(* IEC 61131-3 sources: JingjiangMoonbox/Application/Application/全局, 3 files *)

(* ---- GCL.st ---- *)
(*@CES
Name=GCL
Type=ConstantList
TypeGuid=ffbfa93a-b94d-45fc-a329-229860183b1d
Guid=bcb51df0-81a2-49d0-af31-1b6fd6cdee10
HasDeclaration=True
HasImplementation=False
*)
{DECLARATION}
VAR_GLOBAL CONSTANT
	gc_xUseNewFlyRemove: BOOL:= TRUE;(*新飞点剔除总开关:TRUE=误差平均前用KS_FlyRemove
逐帧剔除并以锁存值替换飞点,FALSE=回退旧飞点判断KS_FB_PickOutFakePoint(旧逻辑完整
保留),改后重新编译生效|Yang.zj+用于新飞点检测 2026.10.24.191149*)
	MASTER_DRIVER_TIME:REAL:= 1;(*运控周期2ms*)
//2026.1.24.215529增加月光宝盒和月光宝盒PRO的类型
	HY_YTPE_CMM_CR_PRO: WORD:= 16#6006;
	HY_YTPE_CMM_CR: WORD:= 16#6005;

	USER_MAX_STATION_NUM_V1:INT:=256;

	gc_iNum_ErrorNum_GT: INT:=3;//gt指令报错执行次数
	gc_iNum_ErrorNum_GT_LOG: INT:=300;//gt指令报错执行次数去写日志
	gc_iTime_s_ServoFailed: INT:=10;//10s伺服打开超时

	gc_lrPi: LREAL:= 3.1415926;
	MAX_UNIT_NUM: INT:=16;(*最大色组数*)
	MAX_STATION_NUM: INT:= 256;
	MAX_AXIS_NUM: INT:= 128;
	(*应对牵引周长算法增加稳速判断等待时长和模拟量滤波计算周长的时长
	默认等待10s和1s调整一次周长*)
	gc_iValueReferToLost: INT:= -32768	;										(*误差标识-丢失|*)
	gc_iValueReferToFakePoint: INT:= -32767	;									(*误差标识-飞点|*)
	gc_iValueReferToSkipTheHeader: INT:= -32766	;							(*误差标识-让料头|*)

	gc_iCycleNum_CalcGirthEvenDelay: INT:= 500;(*算周长算法稳速等待时常，推荐10s(20ms周期就是500个周期)*)
	gc_iCycleNum_CalcDelay: INT:= 500;(*周长计算间隔时长，推荐1s(20ms周期就是50个周期)*)

	gc_tmHold_PreStart				: TIME := T#3S; (* 开机预启动持续时间|该值在程序中赋值给响铃时间| 2022.5.27.143829|该值被弃用*)
	gc_tmHold_PreStart_BeiRen		: TIME := T#6s; (* 北人开机预启动持续时间|和响铃时间是分开的| 2022.5.27.143829*)
	gc_tmAlarmHold_PreStart			: TIME := T#3s; (* 开机预启动报警持续时间| *)
	GC_LRMOTORPPR					: LREAL:=4194304;//2025.7.3.175755
	gc_EXT_TSK_CYCLE_TIME		: INT := 35;(*2023.06.19.102054||niu.j||任务周期35*)
	gc_TENSION_TSK_CYCLE_TIME		: INT := 20;(*2023.06.19.102054||niu.j||任务周期35*)
	gc_MAIN_TSK_CYCLE_TIME		: INT := 10;(*2023.06.19.102054||niu.j||任务周期35*)

	MAX_CMD_NUM_PDU				: INT := 10;(* 最大pdu命令的数量 *)
	MAX_PDU_CMD_BYTES_UP		: INT := 60;(* 来源于1024/16(MAX_UNIT_NUM)/此数必须是4字节的整数倍 *)
	MAX_PDU_CMD_BYTES_DN		: INT := 60;(* 来源于1024/16(MAX_UNIT_NUM)/此数必须是4字节的整数倍 *)
	MAILBOX_PKG_MAX_BYTES		: INT := 480;(* Mailbox包最大长度/2021.11.24.180543/+ *)
	TIMEOUTS_PDU_CMD_CHG		: TIME := T#60MS;(* PDU命令切换超时/2021.12.4.131327/hdp *)
	TIMEOUTS_MAILBOX_FORCESYNC	: TIME := T#100S;(* MAILBOX通讯强制同步超时/2021.12.21.143505/hdp *)

	MAX_KS_UDPPKG_BYTES: UINT := 1024;
	MAX_MEMBLOCK_BYTES: UINT:= (MAX_KS_UDPPKG_BYTES-20);
	PARAM_ZONE_ALTERNATE_OFST: UINT := 0;
	PARAM_ZONE_C2S: UINT := 16384;
	PARAM_ZONE_RESERVED: UINT := 45912;
	REGS_PER_DATA_NODE: UINT := 110;(*每个数据节点的寄存器数量*)
	MAX_DATA_NODE_NUM: UINT := 512;(*最大的数据节点数量*)
	MAX_MB_FIFO_ITEMS: INT := 10;(*ModBus报文FiFo条目上限*)

	CRC_DICTIONARY: ARRAY [0..255] OF WORD :=
		[16#0000, 16#1189, 16#2312, 16#329B, 16#4624, 16#57AD, 16#6536, 16#74BF,
		16#8C48, 16#9DC1, 16#AF5A, 16#BED3, 16#CA6C, 16#DBE5, 16#E97E, 16#F8F7,
		16#1081, 16#0108, 16#3393, 16#221A, 16#56A5, 16#472C, 16#75B7, 16#643E,
		16#9CC9, 16#8D40, 16#BFDB, 16#AE52, 16#DAED, 16#CB64, 16#F9FF, 16#E876,
		16#2102, 16#308B, 16#0210, 16#1399, 16#6726, 16#76AF, 16#4434, 16#55BD,
		16#AD4A, 16#BCC3, 16#8E58, 16#9FD1, 16#EB6E, 16#FAE7, 16#C87C, 16#D9F5,
		16#3183, 16#200A, 16#1291, 16#0318, 16#77A7, 16#662E, 16#54B5, 16#453C,
		16#BDCB, 16#AC42, 16#9ED9, 16#8F50, 16#FBEF, 16#EA66, 16#D8FD, 16#C974,
		16#4204, 16#538D, 16#6116, 16#709F, 16#0420, 16#15A9, 16#2732, 16#36BB,
		16#CE4C, 16#DFC5, 16#ED5E, 16#FCD7, 16#8868, 16#99E1, 16#AB7A, 16#BAF3,
		16#5285, 16#430C, 16#7197, 16#601E, 16#14A1, 16#0528, 16#37B3, 16#263A,
		16#DECD, 16#CF44, 16#FDDF, 16#EC56, 16#98E9, 16#8960, 16#BBFB, 16#AA72,
		16#6306, 16#728F, 16#4014, 16#519D, 16#2522, 16#34AB, 16#0630, 16#17B9,
		16#EF4E, 16#FEC7, 16#CC5C, 16#DDD5, 16#A96A, 16#B8E3, 16#8A78, 16#9BF1,
		16#7387, 16#620E, 16#5095, 16#411C, 16#35A3, 16#242A, 16#16B1, 16#0738,
		16#FFCF, 16#EE46, 16#DCDD, 16#CD54, 16#B9EB, 16#A862, 16#9AF9, 16#8B70,
		16#8408, 16#9581, 16#A71A, 16#B693, 16#C22C, 16#D3A5, 16#E13E, 16#F0B7,
		16#0840, 16#19C9, 16#2B52, 16#3ADB, 16#4E64, 16#5FED, 16#6D76, 16#7CFF,
		16#9489, 16#8500, 16#B79B, 16#A612, 16#D2AD, 16#C324, 16#F1BF, 16#E036,
		16#18C1, 16#0948, 16#3BD3, 16#2A5A, 16#5EE5, 16#4F6C, 16#7DF7, 16#6C7E,
		16#A50A, 16#B483, 16#8618, 16#9791, 16#E32E, 16#F2A7, 16#C03C, 16#D1B5,
		16#2942, 16#38CB, 16#0A50, 16#1BD9, 16#6F66, 16#7EEF, 16#4C74, 16#5DFD,
		16#B58B, 16#A402, 16#9699, 16#8710, 16#F3AF, 16#E226, 16#D0BD, 16#C134,
		16#39C3, 16#284A, 16#1AD1, 16#0B58, 16#7FE7, 16#6E6E, 16#5CF5, 16#4D7C,
		16#C60C, 16#D785, 16#E51E, 16#F497, 16#8028, 16#91A1, 16#A33A, 16#B2B3,
		16#4A44, 16#5BCD, 16#6956, 16#78DF, 16#0C60, 16#1DE9, 16#2F72, 16#3EFB,
		16#D68D, 16#C704, 16#F59F, 16#E416, 16#90A9, 16#8120, 16#B3BB, 16#A232,
		16#5AC5, 16#4B4C, 16#79D7, 16#685E, 16#1CE1, 16#0D68, 16#3FF3, 16#2E7A,
		16#E70E, 16#F687, 16#C41C, 16#D595, 16#A12A, 16#B0A3, 16#8238, 16#93B1,
		16#6B46, 16#7ACF, 16#4854, 16#59DD, 16#2D62, 16#3CEB, 16#0E70, 16#1FF9,
		16#F78F, 16#E606, 16#D49D, 16#C514, 16#B1AB, 16#A022, 16#92B9, 16#8330,
		16#7BC7, 16#6A4E, 16#58D5, 16#495C, 16#3DE3, 16#2C6A, 16#1EF1, 16#0F78];

	(* 通讯信号 *)
	SEMA_UPLOAD					: DWORD := 16#87654321; (* 上行旗语/去主站 *)
	SEMA_DOWNLOAD				: DWORD := 16#12345678; (* 下行旗语/主站来 *)
(*	SEMA_EXT_UPLOAD				: DWORD := 16#56782345; (* 扩展上行旗语/去主站 *)
	SEMA_EXT_DOWNLOAD			: DWORD := 16#23455678; (* 扩展下行旗语/主站来 *)
*)	SEMA_REQ_DISPATCH			: DWORD := 16#51515151; (* 请求旗语/请求主站重新派发指定数据包 *)
	SEMA_PLS_REQ_DISPATCH		: DWORD := 16#A781220A; (* 请非主站重发请求指令(SEMA_REQ_DISPATCH)/主站来 *)
(*	SEMA_SYNC_ING				: DWORD := 16#13572468; (* 状态旗语/正在同步中... *)
	SEMA_SYNC_END				: DWORD := 16#A1A2A3A4; (* 状态旗语/同步完成... *)
*)	SEMA_VIP_COMMAND			: DWORD := 16#19781220; (* 超级旗语/作特殊用途... *)
	SEMA_STANDBY				: DWORD := 16#00000000; (* 复位旗语 *)

	(*2021.7.16.104349 485串口通讯使用|*)
	gc_auchCRCHi:ARRAY [0..255] OF BYTE:=
	[16#00, 16#C1, 16#81, 16#40, 16#01, 16#C0, 16#80, 16#41, 16#01, 16#C0,16#80, 16#41, 16#00, 16#C1, 16#81, 16#40, 16#01, 16#C0, 16#80, 16#41,
	16#00, 16#C1, 16#81, 16#40, 16#00, 16#C1, 16#81, 16#40, 16#01, 16#C0,16#80, 16#41, 16#01, 16#C0, 16#80, 16#41, 16#00, 16#C1, 16#81, 16#40,
	16#00, 16#C1, 16#81, 16#40, 16#01, 16#C0, 16#80, 16#41, 16#00, 16#C1,16#81, 16#40, 16#01, 16#C0, 16#80, 16#41, 16#01, 16#C0, 16#80, 16#41,
	16#00, 16#C1, 16#81, 16#40, 16#01, 16#C0, 16#80, 16#41, 16#00, 16#C1,16#81, 16#40, 16#00, 16#C1, 16#81, 16#40, 16#01, 16#C0, 16#80, 16#41,
	16#00, 16#C1, 16#81, 16#40, 16#01, 16#C0, 16#80, 16#41, 16#01, 16#C0,16#80, 16#41, 16#00, 16#C1, 16#81, 16#40, 16#00, 16#C1, 16#81, 16#40,
	16#01, 16#C0, 16#80, 16#41, 16#01, 16#C0, 16#80, 16#41, 16#00, 16#C1,16#81, 16#40, 16#01, 16#C0, 16#80, 16#41, 16#00, 16#C1, 16#81, 16#40,
	16#00, 16#C1, 16#81, 16#40, 16#01, 16#C0, 16#80, 16#41, 16#01, 16#C0,16#80, 16#41, 16#00, 16#C1, 16#81, 16#40, 16#00, 16#C1, 16#81, 16#40,
	16#01, 16#C0, 16#80, 16#41, 16#00, 16#C1, 16#81, 16#40, 16#01, 16#C0,16#80, 16#41, 16#01, 16#C0, 16#80, 16#41, 16#00, 16#C1, 16#81, 16#40,
	16#00, 16#C1, 16#81, 16#40, 16#01, 16#C0, 16#80, 16#41, 16#01, 16#C0,16#80, 16#41, 16#00, 16#C1, 16#81, 16#40, 16#01, 16#C0, 16#80, 16#41,
	16#00, 16#C1, 16#81, 16#40, 16#00, 16#C1, 16#81, 16#40, 16#01, 16#C0,16#80, 16#41, 16#00, 16#C1, 16#81, 16#40, 16#01, 16#C0, 16#80, 16#41,
	16#01, 16#C0, 16#80, 16#41, 16#00, 16#C1, 16#81, 16#40, 16#01, 16#C0,16#80, 16#41, 16#00, 16#C1, 16#81, 16#40, 16#00, 16#C1, 16#81, 16#40,
	16#01, 16#C0, 16#80, 16#41, 16#01, 16#C0, 16#80, 16#41, 16#00, 16#C1,16#81, 16#40, 16#00, 16#C1, 16#81, 16#40, 16#01, 16#C0, 16#80, 16#41,
	16#00, 16#C1, 16#81, 16#40, 16#01, 16#C0, 16#80, 16#41, 16#01, 16#C0,16#80, 16#41, 16#00, 16#C1, 16#81, 16#40];
	gc_auchCRCLo:ARRAY [0..255] OF BYTE:=
	[16#00, 16#C0, 16#C1, 16#01, 16#C3, 16#03, 16#02, 16#C2, 16#C6, 16#06,16#07, 16#C7, 16#05, 16#C5, 16#C4, 16#04, 16#CC, 16#0C, 16#0D, 16#CD,
	16#0F, 16#CF, 16#CE, 16#0E, 16#0A, 16#CA, 16#CB, 16#0B, 16#C9, 16#09,16#08, 16#C8, 16#D8, 16#18, 16#19, 16#D9, 16#1B, 16#DB, 16#DA, 16#1A,
	16#1E, 16#DE, 16#DF, 16#1F, 16#DD, 16#1D, 16#1C, 16#DC, 16#14, 16#D4,16#D5, 16#15, 16#D7, 16#17, 16#16, 16#D6, 16#D2, 16#12, 16#13, 16#D3,
	16#11, 16#D1, 16#D0, 16#10, 16#F0, 16#30, 16#31, 16#F1, 16#33, 16#F3,16#F2, 16#32, 16#36, 16#F6, 16#F7, 16#37, 16#F5, 16#35, 16#34, 16#F4,
	16#3C, 16#FC, 16#FD, 16#3D, 16#FF, 16#3F, 16#3E, 16#FE, 16#FA, 16#3A,16#3B, 16#FB, 16#39, 16#F9, 16#F8, 16#38, 16#28, 16#E8, 16#E9, 16#29,
	16#EB, 16#2B, 16#2A, 16#EA, 16#EE, 16#2E, 16#2F, 16#EF, 16#2D, 16#ED,16#EC, 16#2C, 16#E4, 16#24, 16#25, 16#E5, 16#27, 16#E7, 16#E6, 16#26,
	16#22, 16#E2, 16#E3, 16#23, 16#E1, 16#21, 16#20, 16#E0, 16#A0, 16#60,16#61, 16#A1, 16#63, 16#A3, 16#A2, 16#62, 16#66, 16#A6, 16#A7, 16#67,
	16#A5, 16#65, 16#64, 16#A4, 16#6C, 16#AC, 16#AD, 16#6D, 16#AF, 16#6F,16#6E, 16#AE, 16#AA, 16#6A, 16#6B, 16#AB, 16#69, 16#A9, 16#A8, 16#68,
	16#78, 16#B8, 16#B9, 16#79, 16#BB, 16#7B, 16#7A, 16#BA, 16#BE, 16#7E,16#7F, 16#BF, 16#7D, 16#BD, 16#BC, 16#7C, 16#B4, 16#74, 16#75, 16#B5,
	16#77, 16#B7, 16#B6, 16#76, 16#72, 16#B2, 16#B3, 16#73, 16#B1, 16#71,16#70, 16#B0, 16#50, 16#90, 16#91, 16#51, 16#93, 16#53, 16#52, 16#92,
	16#96, 16#56, 16#57, 16#97, 16#55, 16#95, 16#94, 16#54, 16#9C, 16#5C,16#5D, 16#9D, 16#5F, 16#9F, 16#9E, 16#5E, 16#5A, 16#9A, 16#9B, 16#5B,
	16#99, 16#59, 16#58, 16#98, 16#88, 16#48, 16#49, 16#89, 16#4B, 16#8B,16#8A, 16#4A, 16#4E, 16#8E, 16#8F, 16#4F, 16#8D, 16#4D, 16#4C, 16#8C,
	16#44, 16#84, 16#85, 16#45, 16#87, 16#47, 16#46, 16#86, 16#82, 16#42,16#43, 16#83, 16#41, 16#81, 16#80, 16#40];
	SEMA_FUNCODE_485_MULT_WR: BYTE:= 16#10;
	SEMA_FUNCODE_485_MULT_RD: BYTE:= 16#03;
	RN_AWR:BYTE:= 16#01;
	RN_ARD:BYTE:= 16#05;

	(* 2025.8.27.154257/han.dp/新合并内容 *)
	FNAME_SYS_CONF: STRING := '/data/kesai/conf/HY.conf';
	FNAME_SYS_PARAM_A: STRING := '/data/kesai/conf/HY-A.bin';
	FNAME_SYS_PARAM_B: STRING := '/data/kesai/conf/HY-B.bin';

(*deprecated@2025.8.27.154330/han.dp
	EACH_MEM_BLOCK_LEN			: DWORD := 4096;(* 每次独立操作的内存块大小 *)
	FILE_BLOCKSIZE_PER_TIMES	: DWORD := 4096;(* 文件操作每次的块大小 *)
	FNAME_SYS_PARAMETERS_A: STRING := '/data/kesai/conf/flexo_A.bin';(* 系统参数文件/2023.8.2.112609/han.dp *)
	FNAME_SYS_PARAMETERS_B: STRING := '/data/kesai/conf/flexo_B.bin';(* 系统参数文件/2023.8.2.112609/han.dp *)
	GC_LOG_ITEM_MAX_NUM							: UINT := 512;(* 日志fifo的最大行数 *)
	(* bit7~bit4/打印信息分类区域/@2021.2.26.111851 *)
	LOG_LEVEL_INFO_NORMAL						: WORD := 16#0080;(* 打印信息/常规 *)
	LOG_LEVEL_INFO_DBG							: WORD := 16#0040;(* 打印信息/程序调试 *)//YY2023.05.20.112732
*)

	gc_byCoatingMaxSum_New			: BYTE := 5; (* 涂布最大轴数-按照列表分配 *)
	gc_dwAbsEnCodeResolution_Uw		: DWORD:=8388608;(*绝对值编码器线束*) (* 2021.8.6.143421/lyt/2^23 *)
	gc_dwAbsEnCodeResolution_Rw		: DWORD:=8388608;(*绝对值编码器线束*) (* 2021.8.6.143421/lyt/2^23 *)

	(*矩阵运算时申请空间所需要的参数|2023.2.16.114926*)
	MATRIX_ROW_MAX:INT:=4;(*矩阵最大行*)
	MATRIX_COLUMN_MAX:INT:=4;(*矩阵最大列*)
	MATRIX_ELEMENT_MAX:INT:=16;(*最大元素|行和列的乘积*)
	//新增运动变量定义|2025.08.05.095813
	GC_LRMOTORPPR_TRAP			:LREAL:=262144.0;//4194304.0;(*Trap电机运动一圈脉冲数*)
	gc_rGirth_Master : REAL := 0.5;
	MAX_ROUNDSAMPLE_NUM: INT:= 4000;(*粗采样点数*)
	gc_iNDEL:INT:=20;(*从压印点到光电眼的幅数*)
	//2025.8.5.101743文件存储
	PREAMBLE: INT := 16#55AA;(* 2023.7.27.110513/han.dp/文件数据桢格式头 *)
	ENDMARK: BYTE := 16#FF;(* 2023.7.27.110513/han.dp/文件数据桢格式尾 *)
	BYTES_PER_ROW_RECORD						: UINT := 8192;(* 每个记录最大的字节数/2021.11.27.150026/hdp *)
	MAX_ROWS_OF_RECORD							: UINT := 5000;(* 记录的最大行/2021.11.27.150411/hdp *)
	PATH_HOME: STRING := '/data/kesai/';
	PATH_HOME_CONF: STRING :='/data/kesai/conf/';
	PATH_HOME_LOG: STRING := '/data/kesai/log/';
	PATH_HOME_DATA: STRING := '/data/kesai/data/';
	MAX_LOG_ITEM_VIEW :INT:= 100 ;
//2025.07.14.160934 | WATCH文件路径
//	PATH_WATCHFILE_1 : STRING := '/opt/codesyscontrol/readCommandTable1.ini';
//	PATH_WATCHFILE_2 : STRING := '/opt/codesyscontrol/readCommandTable2.ini';
//	PATH_WATCHFILE_3 : STRING := '/opt/codesyscontrol/readCommandTable3.ini';
//	PATH_WATCHFILE_4 : STRING := '/opt/codesyscontrol/readCommandTable4.ini';
//	PATH_WATCHFILE_5 : STRING := '/opt/codesyscontrol/readCommandTableEXT.ini';
	PATH_CONFIG_CORE1 : STRING := '/opt/codesyscontrol/gtn_core1.cfg';
	PATH_CONFIG_CORE2 : STRING := '/opt/codesyscontrol/gtn_core2.cfg';
	PATH_WATCHFILE : STRING := '/opt/codesyscontrol/readCommandTable.ini';

	(*2025.8.7.141111*)
	ARC_DELAY_N_MAX:INT:=50;
	ARC_DELAY_N_MAX_DDPD:INT:=200;(*DDPD解耦延时函数缓存大小,"该色到前一色料长/版周长"取整不得大于200*)
	DECOUPLD_DDPD_MAX:INT:=13;(*DDPD共配置13色解耦*)
	DECOUPLD_FDPD_MAX:INT:=13;(*FDPD共配置13色解耦@跟一色隔色解耦*)
	gc_iMaxErrDataItemInList					: INT := 100;(* 误差传递功能的最大存储误差幅数数量 *)
	GC_PU_MAX_NUM								: INT := 16;(* 支持的最大印刷色 *)
	MAX_TSK_CYCLE_MONITORING	: INT := 3;(* 任务周期需要监测的最大数量 *)

(*日志服务新增*)

	GC_LOG_CLASSES_MAX_NUM						: INT := 4;(* 日志种类的数量/[1]总日志/[2]LOG_LEVEL_ALARM/[3]LOG_LEVEL_EVT_/[4]LOG_LEVEL_INFO/ *)

	(* 2021.1.22.163214|为了让过滤更好处理一些|我们从枚举放到了全局常量区域 *)
	(* bit15~bit12/故障报警等分类区域/@2021.2.26.111851 *)
	LOG_LEVEL_ALARM_FATAL						: WORD := 16#8000;(* 致命错误/程序运行都存在问题 *)
	LOG_LEVEL_ALARM_SERIOUS						: WORD := 16#4000;(* 严重报警/会作急停处理 *)
	LOG_LEVEL_ALARM_NORMAL						: WORD := 16#2000;(* 普通报警/不会主动急停 *)
	LOG_LEVEL_ALARM_LOGICCONDITION				: WORD := 16#1000;(* 报警|逻辑条件错误 *)

	(* bit11~bit8/事件记录分类区域/@2021.2.26.111851 *)
	LOG_LEVEL_EVT_USRACTIONS					: WORD := 16#0800;(* 事件记录/用户操作 *)
	LOG_LEVEL_EVT_MOTIONLOGIC					: WORD := 16#0400;(* 事件记录/运动逻辑 *)
	LOG_LEVEL_EVT_PROGRAM_AUTOMATIC				: WORD := 16#0200;(* 事件记录/程序自动触发 *)

	(* bit7~bit4/打印信息分类区域/@2021.2.26.111851 *)

	(* 2023.3.31.091435/han.dp/准备支持日志的部分中文显示 *)
	MAX_ALARMITEM_NUM							: INT := 100;(* 报警条目上限 *)
	(*新增变量-开始|wang.nt|2025.08.13.135942*)
	GC_FORCEDOUT_AXIS_BOUND_L					: INT := 17;(* 强制排除的轴范围左边界从17/最大到GC_PU_MAX_NUM色 *)
	GC_FORCEDOUT_AXIS_BOUND_R					: INT := 20;(* 强制排除的轴范围右边界到20/21开始是B系放料A轴 *)
	(*新增变量-结束|wang.nt|2025.08.13.135942*)

	//2025.08.18.110718 | 增加固高WATCH功能路径
	PATH_HOME_WATCH_DATA: STRING := '/data/kesai/watch/watchData.txt';
 	PATH_HOME_WATCH_CONFIG: STRING := '/opt/codesyscontrol/watchTimer.ini';

	PATH_HOME_WATCH_CONFIG_TEMP: STRING := '/opt/codesyscontrol/watchTimerTemp.ini';

	(*2025.8.19.201228新增*)
	gc_iVirEncPPR: INT:= 8000;

	gc_diVirEncPPR_New			: DINT:= 131072;//131072;//2024.10.23.184529新增的单圈绝对位置累计值 |火眼从65536变换成131072
	//gc_dwMotorPPR								: DWORD := 2097152;(* 电机每转的脉冲数|2^21 *)
	gc_iCycleTime_Motion			: INT := 21; (* 2018.7.1.204007\原始约定| *)
	gc_byInvisCoatingPrnAxisIdx					: BYTE := 20;(* 涂布隐藏轴索引id *)
	gc_byCoatingWay					: BYTE := 5;

//2025.11.24.104500 | 增加修改龙门相关
	gc_iMax_PressureRoller_Unit: INT:=3;//每个色组最大的压力组数
	gc_ResCount_Profile : INT := 64;//单个核的轴资源数
END_VAR
{IMPLEMENTATION}

(* ---- GVL.st ---- *)
(*@CES
Name=GVL
Type=ConstantList
TypeGuid=ffbfa93a-b94d-45fc-a329-229860183b1d
Guid=8a98e878-1566-4378-b3a1-83639989e28b
HasDeclaration=True
HasImplementation=False
*)
{DECLARATION}
VAR_GLOBAL
	g_xRunNormalTask			: BOOL:= FALSE;
	g_iRunStepId				: INT := RUNSTEP_STARTUP;(* 2023.8.3.095049/han.dp *)
	g_xFlag_LogTaskRun			: BOOL;(*文件保存模块运行标志*)
	g_xFlag_OtherTaskRun		: BOOL;(*其他任务*)
	g_xFlag_WriteParamFile		: BOOL;
(*deprecated@2025.8.27.164639/han.dp
	g_stStTravelLogRec: StTravelLogRec;(* 运行日志 *)
*)
	g_stStSts_To_Diamonds_HMI: StParam_Diamonds_Wr;
	g_stStSysParam				: StSysParam;

	(* 2025.8.27.154412/han.dp/合并功能 *)
	g_pstStHYLogFifo			: POINTER TO StHYLogFifo := 0;(* 2025.8.23.170701/han.dp/增加的日志队列 *)
	g_dwMem1MB					: DWORD := 0;(* 2025.8.21.181040/程序进入任务前申请的1M内存 *)
	g_diErrCode_FileProc		: DINT := 0;(* 2025.8.21.181514/文件操作错误代码 *)
	g_pstStUdpOnlySendFifo		: POINTER TO StUdpOnlySendFifo := 0;

(*deprecated@2025.8.27.154430/han.dp
	g_stStSysParam_SaveParam				: StSysParam_SaveParam;
*)

	g_astStAxisRapidAdjProf_V	: ARRAY [1..MAX_UNIT_NUM] OF StAxisRapidAdjProf_V;
	g_astStAxisRapidAdjProf_H	: ARRAY [1..MAX_UNIT_NUM] OF StAxisRapidAdjProf_H;
	g_astStEvtReq				: ARRAY [1..2] OF StEvtReq	;
	g_axCommVel_Sure: ARRAY [1..2,1..3] OF BOOL;(*2019.10.21.095108|常用速度123按钮*)
	g_adiVel_Virtual_Tar: ARRAY [1..2] OF DINT;
	g_alrMax_a_S_pos: ARRAY [1..2] OF LREAL;
	g_alrTime_S: ARRAY [1..2] OF LREAL;
	g_alrJerk_SBegin: ARRAY [1..2] OF LREAL;
	g_alrJerk_SEnd: ARRAY [1..2] OF LREAL;
	g_axMotionEnabled:ARRAY [1..2] OF BOOL;
	g_axis_ctl: INT;
	wTestButton_Input: WORD;
	wTestButton_Output: WORD;
	g_astStIOMap_Main_FE					: ARRAY [1..4] OF StIOMap_Main_FE;(*轴io数据区域|AB系*)
	g_astStIOMap_Axis_FE					: ARRAY [1..MAX_UNIT_NUM] OF StIOMap_Axis_FE;(*轴io数据区域|`````````````````````````````````````````````*)
	g_astStIOMap_Axis_Extra_FE				: ARRAY [1..MAX_UNIT_NUM] OF StIOMap_Axis_Extra_FE;
	g_astStIOMap_UwRw_FE_Uw					: ARRAY [1..2] OF StIOMap_UwRw_FE;(*轴io数据区域|AB系*)
	g_astStIOMap_UwRw_FE_Rw					: ARRAY [1..2] OF StIOMap_UwRw_FE;(*轴io数据区域|AB系*)

//	g_stStRingInfVer1			: StRingInfVer1;
	g_astStSetPrm				: ARRAY [1..MAX_STATION_NUM] OF TSetMultiMcFunctionPrm;
	g_stStGetPrm				: TMultiMcFunctionReadPrm;
	//g_alrVarValue				: ARRAY [1..200] OF LREAL;
	g_astMotionSts 				: ARRAY[1..MAX_STATION_NUM] OF MotionSts;

	g_abyStationList_CommHMI	: ARRAY [1..MAX_STATION_NUM] OF BYTE;
//	g_abyStationList_CommKSCR	: ARRAY [1..MAX_STATION_NUM] OF BYTE;

	(*2025.6.25.211256测试电机运动，完全照搬*)
	g_xStart: BOOL;
	g_mBtn_Init: BOOL;
	g_mBtn_Clr:BOOL:=FALSE;
	g_mBtn_ZeroPos:BOOL:=FALSE;
	g_mBtn_SetMode:BOOL:=FALSE;
	g_mBtn_Start:BOOL:=FALSE;
	g_mBtn_ServerCtl:BOOL:=FALSE;
	g_mBtn_Stop:BOOL:=FALSE;
// 	g_axisId:ARRAY [1..20] OF INT;

// 	g_iAxisId:ARRAY [1..96] OF INT;
// 	g_iServerCtl:BYTE:=0;
// 	core: INT:=1;
// 	g_axisCount:INT:=3;
// 	g_varValue:ARRAY [1..200] OF LREAL;
// 	g_rVel_Cur_HMI_Test:REAL;

	//新增运动相关全局定义|2025.08.05.094744
	//Trap
// 	g_alrTarPos_Horz : ARRAY[1..MAX_UNIT_NUM] OF LREAL := [MAX_UNIT_NUM(1000)];			//um
// 	g_lrMaxVel_Horz : LREAL := 0.2;		//um/ms、mm/s
// 	g_alrTarPos_PhotoCell : ARRAY[1..MAX_UNIT_NUM] OF LREAL := [MAX_UNIT_NUM(10)];			//mm
// 	g_lrMaxVel_PhotoCell : LREAL := 5;
	//Gantry
// 	g_target_pos : LINT := 4194304;
// 	g_max_vel : DINT := 100;
// 	g_diMain : DINT := 0;
// 	g_diSecond : DINT := 0;
	//运动相关
// 	g_astTStTrapParamUser 			: ARRAY[1..MAX_STATION_NUM] OF TStTrapParamUser;
// 	g_astTStJogParamUser 			: ARRAY[1..MAX_STATION_NUM] OF TStJogParamUser;
// 	g_astTStGearParamUser 			: ARRAY[1..MAX_STATION_NUM] OF TStGearParamUser;
// 	g_astTStGantrayTrapParamUser 	: ARRAY[1..MAX_STATION_NUM] OF TStGantrayTrapParamUser;

	g_iAxisNum_Trap					: INT;(*点位运动轴数量*)
	g_aiStationList_Trap			: ARRAY [1..MAX_STATION_NUM] OF INT;(*点位运动轴列表*)
	g_iAxisNum_Gear					: INT;(*电子齿轮运动轴数量*)
	g_aiStationList_Gear			: ARRAY [1..MAX_STATION_NUM] OF INT;(*电子齿轮运动轴列表*)
	g_iAxisNum_GantrayTrap			: INT;(*龙门点位运动组数量*)
	g_aiStationList_GantrayTrap		: ARRAY [1..MAX_STATION_NUM] OF INT;(*龙门点位运动轴列表*)
	g_iAxisNum_Jog					: INT;(*龙门点位运动组数量*)
	g_aiStationList_Jog				: ARRAY [1..MAX_STATION_NUM] OF INT;(*龙门点位运动轴列表*)
	g_iAxisNum_All					: INT;
	g_aiStationList_All				: ARRAY [1..MAX_STATION_NUM] OF INT;
	g_aiIndexList_All_Trap			: ARRAY [1..MAX_STATION_NUM] OF INT;(*点位运动轴列表*)
	g_aiIndexList_All_Gear			: ARRAY [1..MAX_STATION_NUM] OF INT;(*电子齿轮运动轴列表*)
	g_aiIndexList_All_Gantray		: ARRAY [1..MAX_STATION_NUM] OF INT;(*龙门点位运动轴列表*)
	g_aiIndexList_All_Jog			: ARRAY [1..MAX_STATION_NUM] OF INT;(*龙门点位运动轴列表*)

	g_arVel_PrnRoller		: ARRAY[1..2] OF REAL;(* 版辊运行速度*)
	g_arVel_NetRoller		: ARRAY[1..2] of REAL;(* 网辊运行速度*)
	g_arVel_BottomRoller	: ARRAY[1..2] OF REAL;(* 底辊运行速度*)

	g_xFlag_Stop_En_Servo : BOOL;

// 	g_axEn_Motor_Gear : ARRAY [1..2] OF  BOOL;
// 	g_axEn_Motor_Trap :  ARRAY [1..2] OF BOOL;
// 	g_axEn_Motor_Gantry :  ARRAY [1..2] OF BOOL;

	//2025.08.05.094751 | 测试 | 运动控制流程
	g_xInk : BOOL;
	g_xTension : BOOL;
	g_xPrint : BOOL;
	g_xStop : BOOL;
	g_xEstop : BOOL;
	g_xStop_ServoOn:BOOL;
	g_xPreStart : BOOL;
	//g_max_acc:LREAL:=0.4;
	g_lrVel_tar: REAL:= 10;
	g_uiArcAdjValue_Max:UINT:=1000;(*套色调整最大值@1000um|临时做到全局*)
	g_pstStTravelDataRec: POINTER TO StTravelDataRec := 0; (* 实时数据记录缓存 *)
	(*系统时间出错想办法先避免2023.09.12.103011*)
	g_stSysTimedate_Rec: RTS_SYSTIMEDATE;
	g_xInitTime: BOOL;
//	g_stStTravelLogRec: StTravelLogRec;(* 运行日志 *)
(*deprecated@2025.8.27.164745/han.dp
	g_pstStTravelLogRec: POINTER TO StTravelLogRec := 0;
*)
	g_stStTravelDataRec: StTravelDataRec;(* 实时数据记录缓存 *)
(*deprecated@2025.8.27.164827/han.dp
	g_astStTravelLogItem_view: ARRAY [1..GC_LOG_ITEM_MAX_NUM] OF StTravelLogItem;(* 2023.11.23.142330/han.dp/用于查看日志的列表/[1]永远是最新的一条记录 *)
*)
	g_xFileClosed_BecauseEmergency: BOOL := FALSE;(* 由于紧急情况文件关闭的标志 *)
	g_xRst_fileProtect: BOOL := FALSE;
	g_sFilename_datfile: STRING := '';
	g_sFilename_logfile: STRING := '';
	g_iErNo_datfile: INT := 0;
	g_iErNo_logfile: INT := 0;

	g_xSaveFineSampleData :BOOL;//精采样标志
	g_dwPlcLoad :DWORD ; //
	g_astAllAxisErrorTransfer: ARRAY [1..MAX_UNIT_NUM] OF StForArcErrRelay; (* 误差传递使用的队列 *)
	g_pastAllAxisErrorTransfer: POINTER TO ARRAY [1..MAX_UNIT_NUM] OF StForArcErrRelay := 0; (* 误差传递使用的队列 *)
	(*一些占空间比较大的变量|通过allloc获得内存*)
	g_pstStGlobalVarByAllocMem:POINTER TO StGlobalVarByAllocMem;
	g_apbyKp_Arc:ARRAY [1..MAX_UNIT_NUM] OF POINTER TO BYTE;(*套色Kp地址值*)
	g_apbyKi_Arc:ARRAY [1..MAX_UNIT_NUM] OF POINTER TO BYTE;(*套色Ki地址值*)
	g_apbyKd_Arc:ARRAY [1..MAX_UNIT_NUM] OF POINTER TO BYTE;(*套色Kd地址值*)
	g_astStRegAdjMana: ARRAY [1..MAX_UNIT_NUM] OF StRegAdjMana ; (* 套色调整量 *)

	g_astStTaskCycleDetection	: ARRAY [1..MAX_TSK_CYCLE_MONITORING] OF StTaskCycleDetection := [MAX_TSK_CYCLE_MONITORING((xRstDetection:= FALSE, udiCycleCnt:= 0, xCalcIntervalEnabled:= FALSE))];
	g_aiFunctionConsueTime : ARRAY [1..10] OF INT;
	g_iTime_Main_Task : INT;
	g_pstStDatasetARC: POINTER TO StDatasetARC := 0; (* 套色数据记录缓存 *)
//	g_xSaveFineSampleData_ToArc:BOOL;(*保存精采样数据-用于套色保存@通过执行GT_RN_MailWrMultReg函数发送数据到pc机(16#F2)*)
	g_abyActionCtlWay	: ARRAY [1..2] OF BYTE;
	(*新增横向参数-开始|wang.nt|2025.08.09.160741*)
	g_iStepDriveDebugNum: INT := 1; (* 步进电机计算单位脉冲对应的距离的色组号 *)
	g_xStepDriveDebugRun: BOOL; (* 步进电机测试启动 *)
	g_xStepDriveDebugResult_Wr: BOOL; (* 步进电机测试结果写入按钮 *)
	g_diStepDriveDebugPulse: DINT := 60000; (* 测试时输出的脉冲个数；以6000个脉冲一圈 我们默认输出10圈 *)
	g_lrStepDriveDebugPulse_PosAct: LREAL; (* 脉冲完成后位置的变化量 *)
	g_astStDigitalMicroStepDrive: ARRAY [1..MAX_UNIT_NUM] OF StDigitalMicroStepDrive;
	(*横向重复总值*)
	g_abyBtn_HorzPreRegister_Repeat:ARRAY [1..2] OF BYTE;(*重复值的横向按钮@界面使用|=0 不运动|=1 按照轴距离运动|=2 整机按照单个值运动*)
	g_adiPreReg_RepeatVal_H:ARRAY [1..2] OF DINT;
	(*目标值*)
	g_abyBtn_HorzPreRegister_Setup:ARRAY [1..2] OF BYTE;(*目标值的横向按钮@界面使用|=0 不运动|=1 按照轴距离运动|=2 整机按照单个值运动*)
	g_adiPreReg_SetupVal_H:ARRAY [1..2] OF DINT;
	(*新增横向参数-结束|wang.nt|2025.08.09.160741*)

	g_xPressRollerDne_Of_WhenTensionIn:BOOL:=FALSE;(*张力投入时候收牵合压标志|有效表示在张力投入的时候收牵合压并且
											使用牵引使用变频器的时候输出收牵使能*)
	g_xUnPressTop_AllUnPressBtn:BOOL;(*全体离压按钮按下时候方式标志|FALSE=按照延时离压|TRUE=离压到最高处*)
	g_xClearUnPressFlag:BOOL:=FALSE;(*最高点清除离压信号@2023.09.21.141508同步*)
	g_axFlag_PressDne: ARRAY [1..MAX_UNIT_NUM] OF BOOL := [MAX_UNIT_NUM(FALSE)];
	g_arDiamWuCompensate_Uw: ARRAY [1..2] OF REAL;			(*主要用于保存了*)
	g_arDiamWuCompensate_Rw: ARRAY [1..2] OF REAL;			(*主要用于保存了*)
	g_arEstiDia_LowPass_Uw: ARRAY [1..2] OF REAL;			(*主要用于保存了*)
	g_arEstiDia_LowPass_Rw: ARRAY [1..2] OF REAL;			(*主要用于保存了*)
	g_arAntiNotch_Out_Uw: ARRAY [1..2] OF REAL;			(*主要用于保存了*)
	g_arAntiNotch_Out_If: ARRAY [1..2] OF REAL;			(*主要用于保存了*)

	g_astStProgMonitoring						: ARRAY [1..2] OF StProgMonitoring;
	(*新增变量-开始|wang.nt|2025.08.12.162001*)
	g_axKeepAlarm_NoMaterial: ARRAY [1..2] OF BOOL;(*没料持续报警*)
	g_axAlarm_AccOrDecing:ARRAY [1..2] OF BOOL;
	g_axAlarm_CutFinish_Uw:ARRAY [1..2] OF BOOL;
	g_axAlarm_CutFinish_Rw:ARRAY [1..2] OF BOOL;
	g_axAlarm_VolDiamAlarm_Uw:ARRAY [1..2] OF BOOL;
	g_xAlarm_CutDne_Uw: BOOL:=FALSE;(*放料裁切后输出报警标志@时间由界面设置*)
	g_xAtleastOneUnitOverTemp:BOOL;(*至少一色过温标志|用于显示*)
	g_axAxisInchDecing: ARRAY [1..MAX_UNIT_NUM] OF BOOL;(*单运行减速中*)
	(*新增变量-结束|wang.nt|2025.08.12.162001*)
	g_dwNormalWorkRunNum: DWORD;
	g_dwTensionRunNum: DWORD;

	g_iAxisOffCnt_If_OK : INT;
	g_iAxisOffCnt_If_Err : INT;
	(*新增变量-结束|wang.nt|2025.08.12.162001*)
	g_pbyRoundData1: POINTER TO BYTE; (* 存储采样数据T1的波形首地址 *)
	g_pbyRoundData2: POINTER TO BYTE; (* 存储采样数据T2的波形首地址 *)

	(*新增变量-开始|wang.nt|2025.08.13.134901*)
(*deprecated@2025.8.27.165000/han.dp
	g_pstStAlarmLogForView		: POINTER TO StAlarmLogForView := 0;(* 用于存放报警列表内容的 *)
	g_pastStAlarmItemForView	: POINTER TO ARRAY [1..MAX_ALARMITEM_NUM] OF StAlarmItemForView := 0;(* 指向报警显示列表的 *)
*)
	g_abyiNFeedLimitWarnFlag: ARRAY [1..2] OF BYTE;
	g_abyOutFeedLimitWarnFlag: ARRAY [1..2] OF BYTE;
	g_axAlarmHeating:ARRAY [1..2] OF BOOL;(*加热异常报警-用于界面显示*)
	g_xIODebugging: BOOL := FALSE; (* 默认未处于IO测试状态|@2020.11.10.094810 *)
	g_xInTheDiagnosis: BOOL := FALSE; (* 标记当前运行是否在诊断中 *)
	g_dwParaFileImportFailed:DWORD;(*参数导入失败标志|按位标识|.0 1色\.1 2色 依次类推*)
	g_xParaFileExportFailed:BOOL;(*参数导出失败*)
	g_iRtn_CheckFirmWareVer:INT;(*版本检查信息
		-1:参数错误
		\.0:GTSD13版本不一致
		\.1:GTSD16D版本不一致
		\.2:GTSD16M版本不一致
		\.3:GSHD版本不一致*)
	g_xAtleastOneUnitOffline_485:BOOL;(*至少一色485离线*)
	g_xAtleastOneUnitLineBreak_485:BOOL;(*至少一色pt100断线*)
	g_axFlag_Alarm_LD:ARRAY [1..2] OF BOOL;
	g_xAlarm_Rev:BOOL:=FALSE;
	g_iAxisId_Alarm_Rev:INT:=1;
	g_dwAvailPhys_kB:DWORD;
	g_xMemAllocFailed:BOOL;
	g_xEhmiOpened_Master:BOOL;(*主站ehmi未打开*)
	g_xNeedRestartPlc:BOOL;(*需要重启plc*)
	g_axReflectSensorLoss:ARRAY [1..2] OF BOOL;
	g_byAutoBackUpSts:BYTE;(*自动备份状态@=1 提示|=2 显示备份弹窗(强制界面切换到主界面)|PRG_SYNC_UI_UPDATE_\fbKS_FB_GrpFailureProc界面操作或者使用了 *)
(*deprecated@2025.8.27.165059/han.dp
	g_apstStTravelLogRec: ARRAY [1..GC_LOG_CLASSES_MAX_NUM] OF POINTER TO StTravelLogRec; (* 2021.7.5.111146/+/ *)
*)
	(*新增变量-结束|wang.nt|2025.08.13.134919*)
	(*新增工艺相关变量*)
	g_xCoolBlowerOpenByKnob: BOOL := FALSE; (* TRUE:冷风开关旋钮作为打开关闭冷风使能标志|否则为全体冷风打开旋钮打开的色组 *)
	g_xStopCoolBlowerWhenEstop: BOOL := FALSE; (* TRUE:急停停止冷风-- *)
	g_xHotBlowerOpenByKnob: BOOL := FALSE; (* TRUE:热风开关旋钮作为打开关闭热风使能标志|否则为全体热风打开旋钮打开的色组 *)
	g_xStopHotBlowerWhenEstop: BOOL := FALSE; (* TRUE:急停停止热风-- *)
	g_xStopAirExhaustWhenEstop:BOOL:=FALSE;(*TRUE:急停停止排风*)
	g_xUseButton_PreHotBlower:BOOL:=FALSE;(*预热风使用按钮选择*)
	g_xUseButton_PreHeating:BOOL:=FALSE;(*预加热使用按钮选择*)
	g_xflag_printPreHeating:bool:=false;(*印刷开启预加热*)

	//2025.08.18.110718 | 增加固高WATCH功能相关
	g_xWatchOn : BOOL;
	g_xWatchOff : BOOL;
	(*2025.08.20.090543 模块采集的编码器值|未认真处理双收双放结构|2021.4.30.113648*)
	g_dwAbsEncSinglePos_Uw			: DWORD;(*放料编码器单圈值|*)
	g_wAbsEncMultiPos_Uw			: WORD;(*放料料编码器多圈值|*)
	g_dwAbsEncSinglePos_Rw			: DWORD;(*收料编码器单圈值|*)
	g_wAbsEncMultiPos_Rw			: WORD;(*收料料编码器多圈值|*)

	g_byLinkage_Lamp_3_Color:BYTE:=0;(*联动时三色灯颜色|默认=Normal|1=Lost|2=warning@2023.07.07.161402*)
	g_byArcLampDisWay:BYTE:=0;(*三色灯显示模式
							    @0 默认在非印刷的时候按照联动指示用，红色作为急停！
					 			@1 在非印刷的时候不显示三色灯,
								@2 欧诺专用*)
	g_axStartAutoFind: ARRAY [1..2] OF BOOL;(*2023.6.1.161520|分系*)
	g_byTypeStepTest:BYTE;(*阶跃测试类型@=1 横向阶跃|反之纵向阶跃@2023.09.04.230955*)
	g_abyVerManuTrigButton: ARRAY [1..MAX_UNIT_NUM] OF BYTE := [MAX_UNIT_NUM(0)]; (* 纵向手动按钮|转发vs可视化界面操作| =1 向上|=2 向下*)
	g_awVirtualCnt: ARRAY [1..MAX_UNIT_NUM] OF WORD;

	g_aiGrpUnitNum: ARRAY [1..2] OF INT;
	g_aiGrpAxisList: ARRAY [1..2,1..MAX_UNIT_NUM] OF INT; (*系的轴列表*)
	g_aiStepAdj: ARRAY [1..2,1..MAX_UNIT_NUM] OF INT;

	g_axAdjMove_Up : ARRAY [1..MAX_UNIT_NUM] OF BOOL;
	g_axAdjMove_Dn : ARRAY [1..MAX_UNIT_NUM] OF BOOL;
	(*新增绝对值编码器相关*)
	g_stStAbsEncIOModule_Uw : StAbsEncIOModule;
	g_stStAbsEncIOModule_Rw : StAbsEncIOModule;

	g_aiMode_Trap_Rtn : ARRAY [1..MAX_UNIT_NUM] OF INT;
	(*2025.8.22.202521*)

	g_abyClrPrnLenCount: ARRAY [1..2,1..3] OF BYTE := [6(0)]; (* 主界面记米清零点击计数 *)
	g_axClearPrnLen: ARRAY [1..2,1..3] OF BOOL; (* 主界面记米清零按钮 *)(*2020.7.30.111243|记米清零分A/B系|X.^_^*)

	g_xClrSts : BOOL;
	g_iCoreId : INT := 1;
	g_iAxisId : INT := 1;
	(*新增预套准相关变量|wang.nt|2025.08.21.165745*)
	g_axPreRegisterCorrConfirm:ARRAY [1..2] OF BOOL;(*预套准修正量确认|通过印刷自动获得修正量*)
	g_axCorrectConfirmBtnDisplay: ARRAY [1..2] OF BOOL;(*自动获取的预套准修正量确认按钮显示标志*)
	g_iPrewrkSubPageId: INT := 3; (* 预套准子画面id| *)
	g_xLoadRecipe_End: BOOL; (* 读取配方完成标志|用于进行相位回复使能| *)
	g_xReqSaveRecipe: BOOL := FALSE; (* 保存配方按钮 *)
	g_xReqSaveCphRecipe: BOOL;
	g_xReqSaveCphCommonVir: BOOL;
	g_xLoadCphRecipe_End: BOOL;
	g_alrTotalAdjustVal_V:ARRAY [1..MAX_UNIT_NUM] OF LREAL;(*套色总的调整量|用于预套准的修正*)
	g_xFlag_CphCommonVir: BOOL;
	g_xFlag_CphCommonVir_end: BOOL;
	g_xCphaseRestore: BOOL;
	g_xCphaseRestore_end: BOOL;
	(*固定相位保存和读取按钮|2024.6.22.163348*)
	g_axFixedPhaseSave:ARRAY [1..2] OF BOOL;
	g_axFixedPhaseRead:ARRAY [1..2] OF BOOL;
	g_adwIndex: ARRAY [1..2] OF DWORD;

	(*2025.9.5.100111*)
	g_byPseudoRandomSeries				:BYTE:=9;(*伪随机测试级数*)
	g_rPseudoRandomAmplitude			:REAL:=0.03;(*伪随机幅值@m/min\V*)
	(*就直接放初始化里处理吧*)
	g_astStAxisIdListInf: ARRAY [1..128] OF StAxisIdListInf;(*128轴运动控制器所有轴的信息-与cfg文件同步，这样以后的CFG文件可不更改*)
	g_xPseudoRandomEn:BOOL;

	g_xPseudoRandomStart:BOOL;

	g_stStStationInfo_KS	: StStationInfo_KS;(*站列表信息*)
	g_astStStepDriveIOModule: ARRAY [1..MAX_UNIT_NUM] OF StStepDriveIOModule;
	g_astStEnc0410R: ARRAY [1..MAX_UNIT_NUM] OF StEnc0410R;             (* 数组下标代表色组号 *)
	g_abyHorzManuTrigButton: ARRAY [1..MAX_UNIT_NUM] OF BYTE := [MAX_UNIT_NUM(0)]; (* 横向手动按钮|转发vs可视化界面操作| *)
	g_abyHorzManu_HMI				: ARRAY [1..MAX_UNIT_NUM] OF BYTE;
	g_alrGirth_CoatingPrn: ARRAY [1..MAX_UNIT_NUM] OF LREAL; (* 实际用于计算的涂布版周长 *)
	(*2024.01.18.094629 +涂布处理参数*)
	g_stStCoatingAxisInf:StCoatingAxisInf;
	g_alrAI_CoatingHMI: ARRAY [1..MAX_UNIT_NUM] OF LREAL; (* 数组索引代表轴号 *)
	g_axArcErrValid:ARRAY [1..MAX_UNIT_NUM] OF BOOL;
	g_aiArcErr_V:ARRAY [1..MAX_UNIT_NUM] OF INT;(*套色的纵向误差@每圈更新一次并按bit置位表示误差有效*)

	g_axAxisInching: ARRAY [1..MAX_UNIT_NUM] OF BOOL; (* 处于过单运行 *)
//	g_axAxisInchDecing: ARRAY [1..MAX_UNIT_NUM] OF BOOL;(*单运行减速中*)
	g_axAxisInchAccing: ARRAY [1..MAX_UNIT_NUM] OF BOOL;(*单运行加速中*)

	g_auiSendDataCnt_Tcp									:ARRAY [1..8] OF UINT;
	g_auiRecvDataCnt_Tcp									:ARRAY [1..8] OF UINT;
	g_auiRecvErrDataCnt_Tcp								:ARRAY [1..8] OF UINT;
	g_auiTimeOutDataCnt_Tcp								:ARRAY [1..8] OF UINT;
	g_auiSendDataCnt_485									:ARRAY [1..8] OF UINT;
	g_auiRecvDataCnt_485									:ARRAY [1..8] OF UINT;
	g_auiRecvErrDataCnt_485								:ARRAY [1..8] OF UINT;
	g_auiTimeOutDataCnt_485								:ARRAY [1..8] OF UINT;
	g_astStGetMotionSts: ARRAY [1..MAX_STATION_NUM] OF StGetMotionSts;
	g_adiPreRegisterPos: ARRAY [1..MAX_UNIT_NUM] OF DINT;

(*2025.11.1.142853*)
	g_alrMaxVel_PreReg:ARRAY [1..MAX_UNIT_NUM] OF LREAL;//预套准最大速度-时间固定，速度不同

	g_awAxisVirtualCnt: ARRAY [1..MAX_UNIT_NUM] OF WORD; (* 2021.6.25.103841/轴虚拟编码器位置记录/恢复配方后由于重新配置采样会造成轴当前相位清零/用该值先保存恢复之前的位置值 *)
	g_awAxisVirtualSts: ARRAY [1..MAX_UNIT_NUM] OF WORD; (* 2021.6.25.104504/增加的虚拟编码器原始值输入 *)

	g_aiGrpUnitList:ARRAY [1..2,1..MAX_UNIT_NUM] OF INT;(*联动未涂布轴列表|一维数组代表系号|初始值代表隐藏*)

	g_alrVel_VirtualAxis : ARRAY[1..2] OF LREAL;
	g_stStSysCfgStruct: StSysCfgStruct;
	g_xBtn_UpdateSysCfg:  BOOL;(*保存系统配置*)
	g_alrPrfPos : ARRAY [1..MAX_UNIT_NUM] OF LREAL;

	//2025.11.03.103620 | bai.zy | TEST_1103
	(*2021.11.29.142224 同步*)
	(*2020.12.23.211550 增加色组轴在运动过程中停止运动以及停止后加速到目标速度功能|Liu.yt*)
(*	g_xMotionStsSwitchEn:BOOL:=TRUE;(*使用该功能标志*)*)
	g_iMaxVel_StsSwitch:INT:=(*50*)600;(*速度可以切换的最大主机速度值|不要限值-写一个大值*)

	g_abyAxisMotionSts:ARRAY [1..MAX_STATION_NUM] OF BYTE;(*轴运动状态标志|0:同步运动状态.
													  |1:同步运动时停止运动状态.
													  |2:停止运动状态
													  |3:停止运动时加速到单运行速度状态.
													  |4:单运行时减速到停止状态.
													  |5:停止运动时或者使用单运行速度运行时加速到同步运动状态.
													  |6:非同步运动时急停到0状态.
													  |7:非同步运动时空转停机到0状态.*)
	g_axAxisMotionInching:ARRAY [1..MAX_STATION_NUM] OF BOOL;
	g_alrAxisMotionVel:ARRAY [1..MAX_STATION_NUM] OF LREAL;(*轴的速度值*)
	g_axLastAxisMotionInchBtn:ARRAY [1..MAX_STATION_NUM] OF BOOL;
	g_alrAcceleToSync: ARRAY [1..16] OF LREAL:=[16(0.0)];(*用来保证同步的加速度|m/min/ms*)
	g_alrTimeToSync: ARRAY [1..16] OF LREAL;(*用来保证同步的时间|m/min/ms*)
	g_alrRelatePos_Final:ARRAY [1..16,1..16] OF LREAL;(*做成16个轴|
													记录目标轴和当前轴的相对位置值|最后恢复的位置差
													一维下标为当前轴号，二维下标为目标轴号*)
	g_alrRelatePosToSync:ARRAY [1..16,1..16] OF LREAL;(*做成16个轴|
												记录目标轴和当前轴的相对位置值|开始切换到同步状态时的位置差
												一维下标为当前轴号，二维下标为目标轴号*)

	g_axInch : ARRAY [1..MAX_UNIT_NUM] OF BOOL;
	g_axLinkage : ARRAY [1..MAX_UNIT_NUM] OF BOOL;

	g_diSyncErrorLimit : DINT := 83886080;
	g_astStMcgsBtn_HMI: ARRAY [1..MAX_UNIT_NUM] OF StMcgsBtn_HMI;

	g_xInit_StationList:BOOL;

	g_xCutSenSorDelay: BOOL;
//	g_stGT_SystemInfo : GT_SystemInfo;

	g_abyCpu_Load : ARRAY [0..3] OF BYTE;

	g_xFlagEmergencyForFile_tmp : BOOL;

//2025.11.24.104500 | 增加修改龙门相关
	g_astStSetPrm_GantryTrap				: ARRAY [1..MAX_STATION_NUM] OF TSetMultiMcFunctionPrm;

	//压力全体动作
	g_xPressUp_To_Dn : BOOL;//全体合压
	g_xPressDn_To_Up : BOOL;//全体离压
	g_xPressUp_To_Load : BOOL;//全体退出
	g_xPressLoad_To_Up : BOOL;//全体进入
	g_xPressMoveToLoad : BOOL;//换版准备
	g_axFirstMenu : ARRAY [1..5] OF BOOL;
	g_awPressMenu : ARRAY [1..5] OF WORD;

	g_axConfirm:ARRAY [1..3,1..MAX_UNIT_NUM] OF BOOL;

	//增加调试阶段测试压力电机反复来回运行
	g_xPressDebugMode : BOOL;
	g_axPressDebugStart : ARRAY [1..gc_iMax_PressureRoller_Unit,1..MAX_UNIT_NUM] OF BOOL;

	//清除压力电机扭矩保护的标志
	g_xConfirmContinueForward : BOOL;

	g_rPos_press_dn_PrnRoller_Pressure_MM : REAL := 3;

	//
	g_rUp_Dn_Length_MM : ARRAY [1..MAX_UNIT_NUM] OF REAL := [MAX_UNIT_NUM(3)];
//	g_rUp_Dn_Length_MM:REAL:=3;
	g_rPos_press_dn_NetRoller_Pressure_MM : REAL :=3;
	g_xConfirm_Adjust_PressDn : BOOL;

	g_iAxis_Test: INT:= 1;
	g_xTest_MoveFor: BOOL;
	g_xTest_MoveRev: BOOL;
	g_rTest_AllLength: REAL:= 3000;
	g_rTest_StepLength: REAL:= 5;

	g_astStTrapAxisParam_Gantray : ARRAY [1..gc_iMax_PressureRoller_Unit,1..MAX_UNIT_NUM] OF StTrapAxisParam_Gantray;

	g_astStHandWheel: ARRAY[1..MAX_UNIT_NUM] OF StHandWheel;
	g_astStHandWheel_BtnCtl: ARRAY [1..MAX_UNIT_NUM] OF StHandWheel_BtnCtl;
	g_sHandConnectedSignal : STRING;
	g_xModeCalibSwitch : BOOL;
	g_xModeCalibSwitch_Flag : BOOL;

	g_axAuto_Press_Unit: ARRAY [1..MAX_UNIT_NUM] OF BOOL;
	g_axPress_Manu: ARRAY [1..MAX_UNIT_NUM] OF BOOL;
	g_axUnPress_Manu: ARRAY [1..MAX_UNIT_NUM] OF BOOL;

	g_liAbsPos_M : LINT;
	g_liAbsPos_G : LINT;
	g_liAbsPosTrap : LINT;

	//2024.11.22.154437 | bai.zy | 清除压力标定
	g_axResetFlag_FinishCalid : ARRAY [1..MAX_UNIT_NUM] OF BOOL;

	g_astStLatch : ARRAY [1..MAX_UNIT_NUM] OF StLatch;

	g_aliTrapAbsPos :ARRAY [1..MAX_STATION_NUM] OF LINT;
	g_aliM_EncPos :ARRAY [1..MAX_STATION_NUM] OF LINT;

	//检测带长
	g_iSyncBandLen_Unit : INT := 1;
	g_xFlag_AxisInch_Print : BOOL;//整机点动标志

	//2025.03.25.180838 |
	g_rGirthStepBandLen_Kp : REAL := 0.1;
	g_rGirthStepBandLen_Kd : REAL := 0.3;

	//2025.01.23.113618 | 带长检测异常
	g_axCheckBandLenErr : ARRAY [1..MAX_UNIT_NUM] OF BOOL;

	//2025.03.10.171545 | 带长滤波去除极值
	g_xRemoveExtremum : BOOL;

	//2025.02.10.095044 | 增加张力调整方式的开关选择以及增加界面对于新PID调整方式的P、I的输入
	g_xTensionAdjust_NewWay : BOOL;
	g_iTensionAdjust_Kp : INT := 30;
	g_iTensionAdjust_Ki : INT := 60;
	g_xInitPressSlope : BOOL;
	g_rPressValue : REAL := 1000.0;
	g_rPressure_AnalogThreshold : REAL := 0.025;
	//2025.02.10.194406 |
	g_rGirthStep : REAL;//收牵调整量
	g_rGirthStep_Kp : REAL;//收牵调整量
	g_rGirthStep_Ki : REAL;//收牵调整量
	g_lrAnalog_Aver : LREAL;//模拟量平均值
	g_rStep_Compension : REAL;//补偿量
	g_lrCur_PressureValue : LREAL;

	//2025.01.23.085415 | bai.zy | 秦华增加印后牵引的压力传感器
	g_lrTempOF_PrintingOut : LREAL;
	g_lrTempOF : LREAL;

	//交互信号
	g_astStInteraction : ARRAY [1..MAX_UNIT_NUM] OF StInteraction;

	g_stStSysStationInf : StSysStationInf;
	g_stStSysGantryAxisInf : StSysGantryAxisInf;

	//2025.03.19.95021 | 纵向对版标志
// 	g_axArcMoveUp : ARRAY[1..MAX_UNIT_NUM] OF BOOL;
// 	g_axArcMoveDn : ARRAY[1..MAX_UNIT_NUM] OF BOOL;

	//2025.12.27.142247 | + 机器类型，看后面要不要增加到系统参数
	g_iMachineryType : INT;

	g_arTempEncPosBandLength : ARRAY [1..MAX_UNIT_NUM] OF REAL;

	g_axInk_Unit: ARRAY [1..MAX_UNIT_NUM] OF BOOL;

	g_axMoveUp : ARRAY [1..MAX_UNIT_NUM] OF BOOL;
	g_axMoveDn : ARRAY [1..MAX_UNIT_NUM] OF BOOL;
	g_aiTemp : ARRAY [1..8] OF INT := [1,2,3,4,5,6,7,8];

	//2026.01.12.140115 | + | 清除驱动器报警
	g_xClrAlr_HMI : BOOL;

	g_iErrAxisId : INT;
	g_iErrTypeId : INT;
	g_iErrUnitId : INT;
	g_iErrCoreId : INT;

	g_abyInteractionCtl : ARRAY [1..MAX_STATION_NUM] OF BYTE;
	(*2026.01.15.154707//新增品字形柔印机参数-适配版辊垂直移动*)
	g_arFix_RightEdge: ARRAY [1..MAX_UNIT_NUM] OF REAL:=[MAX_UNIT_NUM(120.00)]; //直角边固定机械值 单位:mm 底辊到版辊
	g_arK_TSHAPED_PrnVertical : ARRAY [1..MAX_UNIT_NUM] OF REAL; //比例系数

	//2026.1.28.151219增加GNS本地IO处理
	g_xUseIO_FromGNS_Enable: BOOL;
	g_dwInput_IO_GNS_P6P8: DWORD;
	g_dwInput_IO_GNS_P4P3: DWORD;
	g_dwOutput_IO_GNS_P5P7: DWORD;

	//2026.01.28.114017 | + | 增加横向的位置记忆，此参数需要放在色组的保持参数里面，先放这里吧
	g_aliABSPos_Horiz : ARRAY [1..MAX_UNIT_NUM] OF LINT;
	g_astStSetPrm_Trap				: ARRAY [1..MAX_STATION_NUM] OF TSetMultiMcFunctionPrm;
	g_axLimit_Left_Wr	 					: ARRAY [1..MAX_UNIT_NUM] OF BOOL;//标定横向左右限位值
 	g_axLimit_Right_Wr	 					: ARRAY [1..MAX_UNIT_NUM] OF BOOL;//标定横向左右限位值
	g_axLimit_Left_WrClr	 					: ARRAY [1..MAX_UNIT_NUM] OF BOOL;//清除横向左右标定限位值
 	g_axLimit_Right_WrClr	 					: ARRAY [1..MAX_UNIT_NUM] OF BOOL;//清除横向左右标定限位值

	g_xMoveEnTrap:BOOL:=TRUE;
	g_axMove_Left: ARRAY [1..MAX_UNIT_NUM] OF BOOL;
	g_axMove_Right: ARRAY [1..MAX_UNIT_NUM] OF BOOL;
	g_xInit_TrapPoint: BOOL:= FALSE;
	g_xWashingPrn: BOOL;

	g_xAxis:BOOL;
	g_xjogtest:BOOL;

	//2026.03.14.113537 | + | 增加虚拟码盘异站功能
	(*2022.1.20.103708 增加了虚拟码盘功能需要变量*)
	g_auiSetVirtualEncCfgCnt:ARRAY [1..2] OF UINT;(*异站虚拟码盘参数设置计数*)
	g_xCheckVirtualStsEn:BOOL;(*异站编码器返回状态检查标志|*)
	g_adwVirtualAcrossEnSts:ARRAY [1..2] OF DWORD;(*异站虚拟码盘设置状态返回*)
	g_axVirtualStsChangeFrom2To:ARRAY [1..2] OF BOOL;(*异站虚拟码盘状态由2切换到别的状态标志|有切换对该标志取反切换*)
	g_axReSetEncCfg:ARRAY [1..2] OF BOOL;(*重新设置异站编码器配置*)

	g_aiSetVirtualEnc_ErrCode: ARRAY [1..2] OF INT;
	g_aiVirtualEnc_AxisId_Src: ARRAY [1..2] OF INT;(*虚拟码盘的源轴号*)
	g_aiVirtualEnc_AxisId_Des: ARRAY [1..2] OF INT := [2(1)];(*虚拟码盘的目标轴号*)
	g_aiSetVirtualEncCfgRtn	 : ARRAY [1..2] OF INT;(*虚拟码盘配置返回值*)

	g_StVirtualParam : StVirtualParam;

	g_awAccButton_Count				:ARRAY [1..MAX_UNIT_NUM] OF WORD;
	g_awDecButton_Count			:ARRAY [1..MAX_UNIT_NUM] OF WORD;
	g_awUpAdjButton_Count			:ARRAY [1..MAX_UNIT_NUM] OF WORD;
	g_awDnAdjButton_Count			:ARRAY [1..MAX_UNIT_NUM] OF WORD;
	g_awLeftAdjButton_Count			:ARRAY [1..MAX_UNIT_NUM] OF WORD;
	g_awRightAdjButton_Count			:ARRAY [1..MAX_UNIT_NUM] OF WORD;
	g_awAlarmButton_Count			:ARRAY [1..MAX_UNIT_NUM] OF WORD;

	//2026.1.26.171345 | + | 增加回零位的功能
	g_axBackToHome : ARRAY [1..2] OF BOOL;

	g_aiTestBtn:ARRAY [1..MAX_UNIT_NUM] OF INT;
	g_aiTestBtn1:ARRAY [1..MAX_UNIT_NUM] OF INT;
	g_aiTestBtn2:ARRAY [1..MAX_UNIT_NUM] OF INT;
	g_aiTestBtn3:ARRAY [1..MAX_UNIT_NUM] OF INT;
	g_aiTestBtn4:ARRAY [1..MAX_UNIT_NUM] OF INT;
	g_aiTestBtn5:ARRAY [1..MAX_UNIT_NUM] OF INT;
	g_aiTestBtn6:ARRAY [1..MAX_UNIT_NUM] OF INT;
	g_aiTestBtn7:ARRAY [1..MAX_UNIT_NUM] OF INT;
	g_lrtest:LREAL;
	g_lrtest1:LREAL;
	g_lrtest2:LREAL;
	g_lrtest3:LREAL;
	g_lrtest4:LREAL;
	g_rtest:REAL;
	g_rtest1:REAL;
	g_uitest1:UINT;
	g_uitest2:UINT;

	g_r1test:REAL;
	g_r1test1:REAL;
	g_ui1test1:UINT;
	g_ui1test2:UINT;

	g_lrposM:ARRAY [1..MAX_UNIT_NUM] OF LREAL;
	g_lrposG:ARRAY [1..MAX_UNIT_NUM] OF LREAL;

	g_rposM:ARRAY [1..MAX_UNIT_NUM] OF REAL;
	g_rposG:ARRAY [1..MAX_UNIT_NUM] OF REAL;
	g_uiNum:ARRAY [1..MAX_UNIT_NUM] OF UINT;

	g_alrTrap_EncPos						: ARRAY [1..MAX_UNIT_NUM] OF LREAL;//横向点位轴的规划位置
	g_aiCount_MoveUp						: ARRAY [1..MAX_UNIT_NUM] OF INT;
	g_aiCount_MoveDn						: ARRAY [1..MAX_UNIT_NUM] OF INT;
	g_arStep_Use							: ARRAY [1..MAX_UNIT_NUM] OF REAL;
	g_alrGantryTrapM_EncPos					: ARRAY [1..MAX_UNIT_NUM] OF LREAL;
	g_alrGantryTrapG_EncPos					: ARRAY [1..MAX_UNIT_NUM] OF LREAL;
	g_aiCount_Dn							: ARRAY [1..MAX_UNIT_NUM] OF INT;
	g_aiCount_Up							: ARRAY [1..MAX_UNIT_NUM] OF INT;
	g_aiCount_unLoad						: ARRAY [1..MAX_UNIT_NUM] OF INT;

	g_alrGantryTrap_PrfPos					: ARRAY [1..MAX_UNIT_NUM] OF LREAL;
	g_alrGantryTrapM_PrfPos					: ARRAY [1..MAX_UNIT_NUM] OF LREAL;
	g_alrGantryTrapG_PrfPos					: ARRAY [1..MAX_UNIT_NUM] OF LREAL;
//2026.04.12.171341
	g_alrCurrentAbsPos_Init : ARRAY [1..MAX_STATION_NUM] OF LREAL;
	g_alrCurrentAbsPos_Debug : ARRAY [1..MAX_STATION_NUM] OF LREAL;
	g_alrCurrentAbsPos_Trap : ARRAY [1..MAX_STATION_NUM] OF LREAL;
	g_alrCurrentAbsPos_M : ARRAY [1..MAX_STATION_NUM] OF LREAL;
	g_alrCurrentAbsPos_G : ARRAY [1..MAX_STATION_NUM] OF LREAL;

	g_alrM_EncPos_1u_m : LREAL;
	g_alrM_EncPos_1u_g : LREAL;

	g_astStAxis_Sts_Save_Gear : ARRAY [1..MAX_STATION_NUM] OF StAxis_Sts_Gear;
	g_astStAxis_Sts_Display_Gear : ARRAY [1..MAX_STATION_NUM] OF StAxis_Sts_Gear;
	g_astStAxis_Sts_Save_GantryTrap : ARRAY [1..MAX_STATION_NUM] OF StAxis_Sts_GantryTrap;
	g_astStAxis_Sts_Display_GantryTrap : ARRAY [1..MAX_STATION_NUM] OF StAxis_Sts_GantryTrap;
	g_astStAxis_Sts_Save_Trap : ARRAY [1..MAX_STATION_NUM] OF StAxis_Sts_Trap;
	g_astStAxis_Sts_Display_Trap : ARRAY [1..MAX_STATION_NUM] OF StAxis_Sts_Trap;

//2026.3.2.162241 | 添加用于存储扭矩系数的数组（大小为MAX_STATION_NUM）
	g_arTqCOeff:ARRAY[1..MAX_STATION_NUM] OF REAL;

//2026.05.08.141028 | + | 增加收放料伺服的标志
	g_xUwRwIsServo	: BOOL;

	g_iRtn_MulFunCtl : INT;

	g_adiMasterEven : ARRAY [1..3] OF DINT;
	g_adiSlaveEven : ARRAY [1..3] OF DINT;
	g_adiMasterSlope : ARRAY [1..3] OF DINT;

	//2026.05.09.160415 | + | 增加龙门偏差过大保护
	g_axPressFlag_Stop : ARRAY [1..MAX_UNIT_NUM] OF BOOL;
	g_axBtn_MoveLeft_Horz: ARRAY [1..MAX_UNIT_NUM] OF BOOL;
	g_axBtn_MoveRight_Horz: ARRAY [1..MAX_UNIT_NUM] OF BOOL;
	g_arTrapPos_mm	: ARRAY [1..MAX_UNIT_NUM] OF REAL;

//2026.5.9.181759增加全自动套印一些变量

	g_aiStep_AutoAdjust: ARRAY [1..MAX_UNIT_NUM] OF INT;(*主站全自动套印的找标的执行状态*)
	//g_io_xStartAutoFind:BOOL;
	//xi.hy
	g_astStFiberMoveStepDriver: ARRAY [1..MAX_UNIT_NUM] OF StFiberMoveStepDriver;
	g_xFindMarkCenter:BOOL;
	(* 2022.4.8.203048/hdp (*2026.03.23.163405||粗采样保存wang.xy*)*)
//	g_xSaveRS2file: BOOL := FALSE;
	g_pstStRSampFifo: POINTER TO StRSampFifo := 0;

	g_StiffenTest :BOOL := FALSE;
	g_lrP_Component_Uw:LREAL;
	g_lrI_Component_Uw:LREAL;
	g_lrD_Component_Uw:LREAL;

	g_lrP_Component_Rw:LREAL;
	g_lrI_Component_Rw:LREAL;
	g_lrD_Component_Rw:LREAL;
	(*2026.03.28.182319||wang.xy*)
//	g_rFiberMove:ARRAY [1..2] OF REAL:= [-3,6];//光纤粗调移动距离

//	g_xEnFastPress :BOOL:=TRUE;//当前色找到就合压
	g_xEnFastPress2 :BOOL;//1.5圈直接合压
//	g_xRFailure:BOOL;//粗采样校准失效
//	g_xFFailure:BOOL;//精采样校准失效
	g_EffectiveHumanIntervention:BOOL;//人工干预有效，打开时如果全自动套印三次没找到位置，需要人工干预才能进行下一步
	g_xAllMeanCtl:bool;

	g_xSendResToOnline:BOOL;

	//2026.04.03.233727
	g_rCoffByOnline:REAL:=1/1000;

	//(*2026.04.06.175340||wang.xy全自动套印合压输入*)
	g_axAutoFind_Press:ARRAY [1..MAX_UNIT_NUM] OF BOOL;(*套色Kp地址值*)

//2026.4.11.150854加速度与加加速度
	g_arCur_A: ARRAY [1..2] OF REAL;
	g_arCur_Jerk: ARRAY [1..2] OF REAL;
	g_aiGrpLinkageAxisNum_Pu: ARRAY [1..2] OF INT;
	g_aiGrpLinkageAxisList: ARRAY [1..2,1..MAX_UNIT_NUM] OF INT;

//	g_alrAxisMotionVel:ARRAY [1..MAX_UNIT_NUM] OF LREAL;(*轴的速度值*)

	g_lrPrfVel2 : LREAL;

	g_lrPrfAcc_MasterAxis : LREAL;
	g_alrPrfAcc_MasterAxis2 : ARRAY [1..2] OF LREAL;

	g_lrK:LREAL;
	g_lrB:LREAL;
	g_xLoadParamFild: BOOL:= FALSE;
//2026.4.12.135907为了将裁切放在主任务增加
	g_axSts_Sensor1Ok: ARRAY [1..2] OF BOOL;
	g_axLamp_PreDrive_Debug_Uw: ARRAY [1..2] OF BOOL;
	g_axReqCut_Uw: ARRAY [1..2] OF BOOL;
	g_axTell_KS_PreDrv_CTL_Uw_CuttDne: ARRAY [1..2] OF BOOL;
	//2026.06.02.223725+
	g_axTell_KS_FB_AvoidSomeFilmWithoutAdjust_CuttDne: ARRAY [1..2] OF BOOL;

	//xi.hy新增@七号以后
//	g_astStVarList : ARRAY [1..MAX_STATION_NUM] OF StVarList;

		(*2026.5.7.173444lhy+*)
	g_byOutType:BYTE:=0;(*输出类型@=0 阶跃一定时间|=1 方波输出|=2 伪随机输出@i_xStepBtn有效则接收伪随机量*)
	g_iTestVelSa:INT:=50;(*启动速度m/min*)
//	g_iTestVelSa_ACC:INT:=60;(*加速启动速度m/min*)
//	g_iTestVelSa_DEC:INT:=100;(*减速启动速度m/min*)
	g_uiSquareCycle_ms:UINT:=1000;
	g_uiSquareNum:UINT:=16;(*2026.1.14.192100+方波个数*)
	g_axStepBtn_MotionCtl:ARRAY [1..2] OF BOOL;(*阶跃按钮@外部沿复位*)
	g_arStepVel_MotionCtl:ARRAY [1..2] OF REAL:=[0.03,0.03];(*阶跃速度@m/min*)
	g_auiStepAccDecTime_MotionCtl:ARRAY [1..2] OF UINT:=[0,0];(*加减速时间，简单点使用一个@ms*)
	g_auiStepTotalTime_MotionCtl:ARRAY [1..2] OF UINT:=[16,16];(*输出的总时间@s|默认1s*)
	g_abyStepAxisId_MotionCtl:ARRAY [1..2] OF BYTE:=[3,3];(*阶跃的轴id@默认为非法值*)
	g_axStepping_MotionCtl:ARRAY [1..2] OF BOOL:=[FALSE,FALSE];(*阶跃中标志*)

//2026.5.12.143246|同步超限代码
	g_diVel_Virtual_Tar_Temp : DINT;
	g_lrMax_a_S_pos : LREAL;

	g_axRemoteSetFailed : ARRAY [1..MAX_UNIT_NUM] OF BOOL;
	g_aiCurLabelPos: ARRAY[1..MAX_UNIT_NUM,1..3] OF INT;
    g_arCurLabelWidth: ARRAY[1..MAX_UNIT_NUM,1..3] OF REAL;
    g_rFiberMoveDist: ARRAY[1..MAX_UNIT_NUM,1..2] OF REAL;

//	g_axRemoteSetFailed : ARRAY [1..MAX_UNIT_NUM] OF BOOL;
	g_arRemainDia_Cur: ARRAY [1..2] OF REAL;
	g_xError_SysCfg: BOOL;//系统配置异常
	g_xUnLine_SysStation: BOOL;//网络站点离线
	g_xTrigSave_BlackoutSts: BOOL;
//2026.05.23.111030 | + |相位恢复超时报警标志
	g_axPhaseRestore_Overtime:  ARRAY [1..2] OF BOOL;
(*2026.5.28.150112增加预套准结构初始化*)
	g_pstStMechanicalParam_01: POINTER TO StMechanicalParam_01; (* 机械结构1 *)
	g_pstStMechanicalParam_02: POINTER TO StMechanicalParam_02; (* 机械结构2 *)
	g_pstStMechanicalParam_03: POINTER TO StMechanicalParam_03; (* 机械结构3 *)
	(*2023.09.21.145817 同步*)
	g_pstStMechanicalParam_05: POINTER TO StMechanicalParam_05;(*机械结构5|2023.07.11.110800*)
//2026.5.29.153619
	g_xAutoPrintMasterAlarm : ARRAY [1..2] OF BOOL;

END_VAR
{IMPLEMENTATION}

(* ---- VER.st ---- *)
(*@CES
Name=VER
Type=ConstantList
TypeGuid=ffbfa93a-b94d-45fc-a329-229860183b1d
Guid=5d11c678-8099-465f-ae42-1f896e770119
HasDeclaration=True
HasImplementation=False
*)
{DECLARATION}
VAR_GLOBAL
//	gc_sVersion: STRING:= '2025.7.3.102405';
//	gc_sVersion: STRING:= '2025.7.4.214233';
	(*合并金刚通讯*)
//	gc_sVersion: STRING:= 'KSFieryEyes-MASTER_V1.0.1-2025.8.26.144842';
	(*更新速度计算对应关系
	更新lib库，增加相机拍照减速比设置
	*)
	(*2025.8.5.200223|更新金刚通讯前备份了一下8.5版本*)
	(*2025.8.6.175048|增加金刚界面参数赋值及参数保存、套色调整算法|niuj*)

	(*v1.0.1版本更新内容：
		1）主站与金刚通讯结构体更新
		2）天枢粗采样数据读取-保存待加
		3）S曲线规划
		4）套色调整
		5）时间：2025.8.26.145356*)
(*	gc_sVersion: STRING:= 'KSFieryEyes-MASTER_V1.0.2-2025.8.27.152843';*)
	(*合并韩工最新关于日志和数据保存相关改动2025.8.27.152907*)
(*	gc_sVersion: STRING:= 'KSFieryEyes-MASTER_V1.0.2-2025.9.6.104807';*)
	(*调整完全放在同一个任务里把2025.9.1.201639*)
(*	gc_sVersion: STRING:= 'KSFieryEyes-MASTER_V1.0.2-2025.9.8.094600';*)
	(*测试完伪随机和增加读取站列表内容*)
(*	gc_sVersion: STRING:= 'KSFieryEyes-MASTER_V1.0.2-2025.9.10.193907';*)
(*横向调整代码和IO输入输出全部放到主任务*)
(*通讯任务更改为10ms*)
(*	gc_sVersion: STRING:= 'KSFieryEyes-MASTER_V1.0.2-2025.9.12.192152';*)
(*出差前最后版本2025.9.12.192201*)
//	gc_sVersion: STRING:= 'KSFieryEyes-MASTER_V1.0.2-2025.9.18.142623';
(*第一次印刷后版本更新|
验证套色调整输出
张力算法
界面伪随机相关变量增加

*)
(*	gc_sVersion: STRING:= 'KSFieryEyes-MASTER_V1.0.2-2025.11.1.164946';*)
(*
1.更新润新发现的一些问题
2.运动功能标准化
3.单运行、预套准
4.系统配置等金刚通讯
*)
(*	gc_sVersion: STRING:= 'KSFieryEyes-MASTER_V1.0.2-2025.11.14.093524';

运城制版测试
*)
(*	gc_sVersion: STRING:= 'KSFieryEyes-MASTER_V1.0.2-2025.11.15.165030';
增加低通滤波频率下发*)
(*	gc_sVersion: STRING:= 'KSFieryEyes-MASTER_V1.0.2-2025.11.16.112443';*)
(*增加获取CPU和内存大小，修改解耦相关内容*)
	//gc_sVersion: STRING:= 'KSFieryEyes-MASTER_V1.0.2-2025.12.30.164122';
(*2025.12.30.164126
1.增加牵引变频控制
2.秦华逻辑增加
3.统一拓扑图
*)
//	gc_sVersion: STRING:= 'KSFieryEyes-MASTER_V1.0.6-2026.03.16.171137';
//2026.03.11.093012 | + | 同步获取编码器位数和最大转速的功能 下面的这一段改成自动的，不使用强制了，已经在秦华验证过
//2026.03.09.170159 | + |一色压辊自动处理
//2026.03.11.100402 | + | 使用Bit26作为压力电机自动合压开关
//2026.03.11.103736 | + | 停机维持伺服、停机上下伺服
//2026.03.12.102825 | + | 同步天枢的数据存储开关
//2026.03.14.113537 | + | 增加虚拟码盘异站功能
//2026.03.16.141753 | + | 增加日志打印
//2026.03.16.171137 | + | 增加单运行方向判断

//gc_sVersion: STRING:= 'KSFieryEyes-MASTER_V1.0.7-2026.03.27.175514';
//2026.03.27.175514 | + | 给超旭同步秦华的金刚清除报警功能    2026.1.27.141112 | + | 增加清除报警的功能

//gc_sVersion: STRING:= 'KSFieryEyes-MASTER_V1.0.10-2026.5.15.115700';
//gc_sVersion: STRING:= 'KSFieryEyes-MASTER_V1.0.11-2026.5.16.112818';
//2026.5.16.112820更新内容
(*
1.预套准参数保存失败原因：预套准结构变量输入写死，更新为变量
2.卷径检测界面变量绑定问题，输入问题；需同步更新金刚界面，
*)
//gc_sVersion: STRING:= 'KSFieryEyes-MASTER_V1.0.11-2026.5.20.091328';
//实时同步程序
(*
1.修复裁切问题
2.修复套色不调整问题
3.修复配方恢复问题
4.更新轴运动状态监控变量表
*)
//gc_sVersion: STRING:= 'KSFieryEyes-MASTER_V1.0.11-2026.5.30.112337';
//gc_sVersion: STRING:= 'KSFieryEyes-MASTER_V1.0.11-2026.07.30.103148';
(*
近期更新：
1.色组控制轴保存数据的枚举位置
2.配方使用的bug,无法写入
3.刮刀手动频率功能块的赋值
4.保存系统配置的同步
5.横向伺服当前位置改为单向通讯
6.主从双向通讯删除了部分按钮计数
7.增加电压实时值和设定值的金刚通讯
8.更新了光纤行走基准定位功能bug
9.更新了xAxisBLocaltion_Out变量书写错误
10.横向伺服当前位置改为单向通讯删除时，没有保留位置，导致通讯有问题
11.增加横向预套准功能输出
12.增加停机时联动轴维持使能功能
*)
//gc_sVersion: STRING:= 'KSFieryEyes-MASTER_V1.0.11-2026.08.19.102507';
(*
绍兴程序独立迭代
1.修复从站停止按钮不清除
2.收放料变频器报警输入
*)
//gc_sVersion: STRING:= 'KSFieryEyes-MASTER_V1.0.11-2026.08.21.132221';
(*
1.增加涂布功能
2.屏蔽报警功能块收放料变频器报警的输入并且保存报警的点位pstStRecord_T^.wPreHotRollerFrq
*)
//gc_sVersion: STRING:= 'KSFieryEyes-MASTER_V1.0.11-2026.08.25.162455';
(*
2026.08.25.143216+使用料膜厚度rFilmThickNess_Using的默认值改为0.02
2026.08.25.143222+收料接料后的预估卷径方向rDiaPrf_CutDne反了，应该是加
*)
//gc_sVersion: STRING:= 'KSFieryEyes-MASTER_V1.0.11-2026.09.02.090905';
(*
2026.09.02.090923+05结构预套准更新
*)
//gc_sVersion: STRING:= 'KSFieryEyes-MASTER_V1.0.11-2026.09.04.142650';
(*
2026.09.04.142708+更新行走机构控制@和欧诺第二台一致
2026.09.04.142724+修复异站功能块bug
2026.09.06.104859+非停机状态下，版辊单运行标志的清除 并且 增加设备类型等于4时，联动色组不允许单运行
*)
//gc_sVersion: STRING:= 'KSFieryEyes-MASTER_V1.0.12-2026.09.12.170702';
(*
2026.09.12.170716+预套准机械参数之后预留120字节
*)
gc_sVersion: STRING:= 'KSFieryEyes-MASTER_V1.0.12-2026.09.13.133606';
(*
2026.09.13.133619| + |增加获取虚拟码盘时返回值错误之后的保护
*)
END_VAR
{IMPLEMENTATION}
